// TIA Portal V20 export
FUNCTION_BLOCK "06_Grundstellungen"   // FB114, FBD
{ S7_Optimized_Access := 'TRUE' }
// stored: MemoryReserve 100, SetENOAutomatically false
   VAR_TEMP
      StörungDW : Int;
      Achse31_GS : Bool;
      GS_Z_Achse1 : Bool;
      GS_Z_Achse2 : Bool;
      GS_Z_Achse3 : Bool;
      GS_Z_Achse4 : Bool;
      GS_Schlitten_POS9_3 : Bool;
   END_VAR
BEGIN

NETWORK
TITLE = Grundstellung gesamt
      A     "Global_Signal"."M_Grundstellung_POS3.0";

      AN    "ProDiag_Allgemein_DB".State.All;
      =     "HMI_COM".Grundstellung_Gesamt;

NETWORK
TITLE = Grundstellung POS3.0
      AN    "POS3_0_Prodiag_DB".State.C1;
      A(;
      O     "POS3_0_Signal"."-1001T1 Oriental_Positionen".POS_OK_Position[0];
      O     "POS3_0_Signal"."-1001T1 Oriental_Positionen".POS_OK_Position[1];
      );
      A(;
      O     "POS3_0_Signal"."-1002T1 Oriental_Positionen".POS_OK_Position[0];
      O     "POS3_0_Signal"."-1002T1 Oriental_Positionen".POS_OK_Position[1];
      );
      AN    "POS3_0_Signal".Station.SK_Richten_gestartet;
      =     "Global_Signal"."M_Grundstellung_POS3.0";


NETWORK
TITLE = Station Sicher Pos3.0
      AN    "POS3_0_Prodiag_DB".State.C1;

      =     "HMI_BETR_ART_POS".POS3_0.Status_Sicher;

END_FUNCTION_BLOCK
